// TIA Portal V21 export
// export: Created 2026-11-11T00:47:28.2882163Z, ExportSetting WithDefaults, DisplayName Totally Integrated Automation Portal, DisplayVersion V21 Update 3, DisplayName STEP 7 Professional, DisplayVersion V21 Update 3, DisplayName STEP 7 Safety, DisplayVersion V21, DisplayName Tech WebApplication, DisplayVersion V21, DisplayName WinCC Basic/Comfort/Advanced, DisplayVersion V21 Update 3, DisplayName WinCC Unified, DisplayVersion V21 Update 3
FUNCTION_BLOCK "FB_Fbd_ex109"   // FB121, FBD
{ S7_Optimized_Access := 'TRUE' }
VERSION : 0.1
// stored: AutoNumber true, IsIECCheckEnabled false, IsRetainMemResEnabled false, MemoryReserve 100, SetENOAutomatically false, UDAEnableTagReadback false
   VAR_INPUT
      v_ob_nr : Int;
      v_dtime : Time;
      v_sign : Word;
   END_VAR
   VAR_OUTPUT
      v_ret_val : Int;
   END_VAR
BEGIN

REGION Network 1: SRT_DINT - Start time-delay interrupt
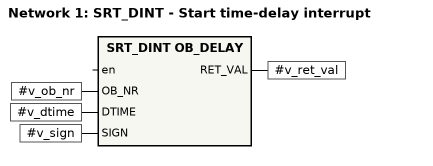
   #v_ret_val := SRT_DINT(OB_NR := #v_ob_nr, DTIME := #v_dtime, SIGN := #v_sign);
END_REGION
END_FUNCTION_BLOCK
